  movel([-0.240083, -0.819456, -2.773882, -1.119051, 1.570796, 1.330713],accel_mss,speed_ms,0,blend_radius_m)
  movel([-0.246972, -0.827519, -2.772360, -1.112509, 1.570796, 1.323824],accel_mss,speed_ms,0,blend_radius_m)
  movel([-0.253406, -0.835845, -2.770751, -1.105793, 1.570796, 1.317390],accel_mss,speed_ms,0,blend_radius_m)
  movel([-0.259324, -0.844374, -2.769062, -1.098952, 1.570796, 1.311472],accel_mss,speed_ms,0,blend_radius_m)
  movel([-0.264353, -0.852401, -2.767435, -1.092553, 1.570796, 1.306443],accel_mss,speed_ms,0,blend_radius_m)
  movel([-0.268744, -0.860169, -2.765824, -1.086396, 1.570796, 1.302052],accel_mss,speed_ms,0,blend_radius_m)
  movel([-0.272465, -0.867667, -2.764235, -1.080487, 1.570796, 1.298331],accel_mss,speed_ms,0,blend_radius_m)
  movel([-0.275488, -0.874892, -2.762673, -1.074824, 1.570796, 1.295308],accel_mss,speed_ms,0,blend_radius_m)
  movel([-0.276730, -0.878403, -2.761902, -1.072084, 1.570796, 1.294066],accel_mss,speed_ms,0,blend_radius_m)
  movel([-0.278648, -0.885206, -2.760387, -1.066796, 1.570796, 1.292148],accel_mss,speed_ms,0,blend_radius_m)
  movel([-0.279316, -0.888500, -2.759643, -1.064245, 1.570796, 1.291480],accel_mss,speed_ms,0,blend_radius_m)
  movel([-0.280060, -0.894869, -2.758187, -1.059334, 1.570796, 1.290737],accel_mss,speed_ms,0,blend_radius_m)
  movel([-0.280127, -0.897947, -2.757473, -1.056968, 1.570796, 1.290669],accel_mss,speed_ms,0,blend_radius_m)
  movel([-0.279987, -0.900948, -2.756772, -1.054668, 1.570796, 1.290809],accel_mss,speed_ms,0,blend_radius_m)
  movel([-0.279491, -0.905065, -2.755801, -1.051523, 1.570796, 1.291305],accel_mss,speed_ms,0,blend_radius_m)
  movel([-0.278705, -0.908998, -2.754863, -1.048528, 1.570796, 1.292092],accel_mss,speed_ms,0,blend_radius_m)
  movel([-0.277654, -0.912736, -2.753962, -1.045690, 1.570796, 1.293142],accel_mss,speed_ms,0,blend_radius_m)
  movel([-0.276370, -0.916287, -2.753099, -1.043004, 1.570796, 1.294426],accel_mss,speed_ms,0,blend_radius_m)
  movel([-0.274870, -0.919629, -2.752278, -1.040482, 1.570796, 1.295926],accel_mss,speed_ms,0,blend_radius_m)
  movel([-0.273177, -0.922754, -2.751504, -1.038131, 1.570796, 1.297619],accel_mss,speed_ms,0,blend_radius_m)
  movel([-0.271316, -0.925662, -2.750778, -1.035949, 1.570796, 1.299480],accel_mss,speed_ms,0,blend_radius_m)
  movel([-0.269306, -0.928336, -2.750106, -1.033947, 1.570796, 1.301490],accel_mss,speed_ms,0,blend_radius_m)
  movel([-0.260160, -0.937511, -2.747762, -1.027116, 1.570796, 1.310636],accel_mss,speed_ms,0,blend_radius_m)
  movel([-0.253034, -0.945065, -2.745789, -1.021535, 1.570796, 1.317763],accel_mss,speed_ms,0,blend_radius_m)
  movel([-0.252477, -0.945898, -2.745569, -1.020921, 1.570796, 1.318320],accel_mss,speed_ms,0,blend_radius_m)
  movel([-0.246274, -0.937106, -2.747867, -1.027417, 1.570796, 1.324523],accel_mss,speed_ms,0,blend_radius_m)
  movel([-0.239566, -0.928371, -2.750097, -1.033921, 1.570796, 1.331230],accel_mss,speed_ms,0,blend_radius_m)
  movel([-0.232400, -0.919726, -2.752254, -1.040409, 1.570796, 1.338397],accel_mss,speed_ms,0,blend_radius_m)
  movel([-0.224833, -0.911212, -2.754331, -1.046846, 1.570796, 1.345963],accel_mss,speed_ms,0,blend_radius_m)
  movel([-0.216924, -0.902878, -2.756318, -1.053193, 1.570796, 1.353873],accel_mss,speed_ms,0,blend_radius_m)
  movel([-0.208734, -0.894762, -2.758211, -1.059416, 1.570796, 1.362062],accel_mss,speed_ms,0,blend_radius_m)
  movel([-0.200327, -0.886916, -2.760002, -1.065471, 1.570796, 1.370469],accel_mss,speed_ms,0,blend_radius_m)
  movel([-0.191774, -0.879388, -2.761684, -1.071317, 1.570796, 1.379022],accel_mss,speed_ms,0,blend_radius_m)
  movel([-0.187679, -0.876001, -2.762430, -1.073958, 1.570796, 1.383118],accel_mss,speed_ms,0,blend_radius_m)
  movel([-0.183450, -0.872734, -2.763143, -1.076512, 1.570796, 1.387346],accel_mss,speed_ms,0,blend_radius_m)
  movel([-0.179125, -0.869625, -2.763815, -1.078949, 1.570796, 1.391671],accel_mss,speed_ms,0,blend_radius_m)
  movel([-0.174747, -0.866715, -2.764439, -1.081235, 1.570796, 1.396049],accel_mss,speed_ms,0,blend_radius_m)
  movel([-0.170354, -0.864043, -2.765007, -1.083339, 1.570796, 1.400443],accel_mss,speed_ms,0,blend_radius_m)
  movel([-0.165982, -0.861648, -2.765513, -1.085228, 1.570796, 1.404814],accel_mss,speed_ms,0,blend_radius_m)
  movel([-0.161676, -0.859568, -2.765950, -1.086871, 1.570796, 1.409121],accel_mss,speed_ms,0,blend_radius_m)
  movel([-0.157477, -0.857842, -2.766310, -1.088237, 1.570796, 1.413319],accel_mss,speed_ms,0,blend_radius_m)
  movel([-0.153425, -0.856510, -2.766587, -1.089292, 1.570796, 1.417371],accel_mss,speed_ms,0,blend_radius_m)
  movel([-0.149560, -0.855608, -2.766774, -1.090007, 1.570796, 1.421237],accel_mss,speed_ms,0,blend_radius_m)
  movel([-0.145927, -0.855177, -2.766863, -1.090349, 1.570796, 1.424869],accel_mss,speed_ms,0,blend_radius_m)
  movel([-0.142567, -0.855251, -2.766848, -1.090290, 1.570796, 1.428229],accel_mss,speed_ms,0,blend_radius_m)
  movel([-0.139522, -0.855865, -2.766721, -1.089803, 1.570796, 1.431274],accel_mss,speed_ms,0,blend_radius_m)
  movel([-0.136824, -0.857050, -2.766475, -1.088864, 1.570796, 1.433972],accel_mss,speed_ms,0,blend_radius_m)
  movel([-0.134519, -0.858837, -2.766102, -1.087449, 1.570796, 1.436278],accel_mss,speed_ms,0,blend_radius_m)
  movel([-0.132645, -0.861261, -2.765595, -1.085534, 1.570796, 1.438152],accel_mss,speed_ms,0,blend_radius_m)
  movel([-0.130842, -0.865165, -2.764769, -1.082455, 1.570796, 1.439954],accel_mss,speed_ms,0,blend_radius_m)
  movel([-0.129631, -0.869711, -2.763796, -1.078881, 1.570796, 1.441165],accel_mss,speed_ms,0,blend_radius_m)
  movel([-0.128936, -0.874759, -2.762702, -1.074928, 1.570796, 1.441860],accel_mss,speed_ms,0,blend_radius_m)
  movel([-0.128670, -0.880175, -2.761510, -1.070704, 1.570796, 1.442126],accel_mss,speed_ms,0,blend_radius_m)
  movel([-0.128760, -0.885825, -2.760248, -1.066316, 1.570796, 1.442036],accel_mss,speed_ms,0,blend_radius_m)
  movel([-0.129131, -0.891586, -2.758941, -1.061862, 1.570796, 1.441665],accel_mss,speed_ms,0,blend_radius_m)
  movel([-0.130394, -0.902931, -2.756306, -1.053152, 1.570796, 1.440402],accel_mss,speed_ms,0,blend_radius_m)
  movel([-0.131557, -0.910187, -2.754578, -1.047624, 1.570796, 1.439239],accel_mss,speed_ms,0,blend_radius_m)
  movel([-0.133085, -0.917458, -2.752812, -1.042119, 1.570796, 1.437712],accel_mss,speed_ms,0,blend_radius_m)
  movel([-0.134926, -0.924737, -2.751010, -1.036643, 1.570796, 1.435870],accel_mss,speed_ms,0,blend_radius_m)
  movel([-0.137037, -0.932034, -2.749168, -1.031187, 1.570796, 1.433760],accel_mss,speed_ms,0,blend_radius_m)
  movel([-0.139370, -0.939343, -2.747287, -1.025759, 1.570796, 1.431427],accel_mss,speed_ms,0,blend_radius_m)
  movel([-0.141879, -0.946667, -2.745366, -1.020356, 1.570796, 1.428917],accel_mss,speed_ms,0,blend_radius_m)
  movel([-0.147269, -0.961389, -2.741392, -1.009608, 1.570796, 1.423527],accel_mss,speed_ms,0,blend_radius_m)
  movel([-0.140519, -0.960936, -2.741517, -1.009936, 1.570796, 1.430278],accel_mss,speed_ms,0,blend_radius_m)
  movel([-0.137016, -0.960927, -2.741519, -1.009943, 1.570796, 1.433781],accel_mss,speed_ms,0,blend_radius_m)
  movel([-0.133979, -0.961411, -2.741386, -1.009592, 1.570796, 1.436818],accel_mss,speed_ms,0,blend_radius_m)
  movel([-0.132765, -0.961921, -2.741245, -1.009222, 1.570796, 1.438031],accel_mss,speed_ms,0,blend_radius_m)
  movel([-0.131825, -0.962655, -2.741043, -1.008690, 1.570796, 1.438971],accel_mss,speed_ms,0,blend_radius_m)
  movel([-0.131206, -0.963639, -2.740771, -1.007979, 1.570796, 1.439590],accel_mss,speed_ms,0,blend_radius_m)
  movel([-0.130958, -0.964905, -2.740420, -1.007064, 1.570796, 1.439839],accel_mss,speed_ms,0,blend_radius_m)
  movel([-0.131131, -0.966478, -2.739983, -1.005928, 1.570796, 1.439665],accel_mss,speed_ms,0,blend_radius_m)
  movel([-0.131778, -0.968398, -2.739446, -1.004544, 1.570796, 1.439018],accel_mss,speed_ms,0,blend_radius_m)
  movel([-0.132943, -0.970690, -2.738802, -1.002896, 1.570796, 1.437853],accel_mss,speed_ms,0,blend_radius_m)
  movel([-0.134674, -0.973378, -2.738043, -1.000969, 1.570796, 1.436123],accel_mss,speed_ms,0,blend_radius_m)
  movel([-0.136314, -0.975590, -2.737413, -0.999386, 1.570796, 1.434482],accel_mss,speed_ms,0,blend_radius_m)
  movel([-0.137990, -0.977600, -2.736838, -0.997950, 1.570796, 1.432806],accel_mss,speed_ms,0,blend_radius_m)
  movel([-0.139696, -0.979424, -2.736314, -0.996651, 1.570796, 1.431100],accel_mss,speed_ms,0,blend_radius_m)
  movel([-0.143196, -0.982582, -2.735401, -0.994406, 1.570796, 1.427601],accel_mss,speed_ms,0,blend_radius_m)
  movel([-0.144982, -0.983947, -2.735004, -0.993438, 1.570796, 1.425815],accel_mss,speed_ms,0,blend_radius_m)
  movel([-0.148619, -0.986335, -2.734306, -0.991748, 1.570796, 1.422177],accel_mss,speed_ms,0,blend_radius_m)
  movel([-0.152315, -0.988361, -2.733710, -0.990318, 1.570796, 1.418481],accel_mss,speed_ms,0,blend_radius_m)
  movel([-0.156050, -0.990151, -2.733182, -0.989056, 1.570796, 1.414746],accel_mss,speed_ms,0,blend_radius_m)
  movel([-0.163527, -0.993487, -2.732190, -0.986712, 1.570796, 1.407269],accel_mss,speed_ms,0,blend_radius_m)
  movel([-0.166909, -0.999532, -2.730372, -0.982486, 1.570796, 1.403888],accel_mss,speed_ms,0,blend_radius_m)
  movel([-0.168793, -1.002571, -2.729447, -0.980371, 1.570796, 1.402004],accel_mss,speed_ms,0,blend_radius_m)
  movel([-0.170824, -1.005546, -2.728535, -0.978308, 1.570796, 1.399972],accel_mss,speed_ms,0,blend_radius_m)
  movel([-0.173015, -1.008396, -2.727655, -0.976338, 1.570796, 1.397781],accel_mss,speed_ms,0,blend_radius_m)
  movel([-0.175376, -1.011062, -2.726826, -0.974501, 1.570796, 1.395420],accel_mss,speed_ms,0,blend_radius_m)
  movel([-0.177921, -1.013486, -2.726068, -0.972835, 1.570796, 1.392875],accel_mss,speed_ms,0,blend_radius_m)
  movel([-0.180668, -1.015618, -2.725397, -0.971375, 1.570796, 1.390128],accel_mss,speed_ms,0,blend_radius_m)
  movel([-0.182641, -1.016748, -2.725040, -0.970601, 1.570796, 1.388155],accel_mss,speed_ms,0,blend_radius_m)
  movel([-0.184252, -1.017225, -2.724889, -0.970275, 1.570796, 1.386545],accel_mss,speed_ms,0,blend_radius_m)
  movel([-0.185536, -1.017141, -2.724915, -0.970332, 1.570796, 1.385261],accel_mss,speed_ms,0,blend_radius_m)
  movel([-0.186525, -1.016588, -2.725090, -0.970711, 1.570796, 1.384271],accel_mss,speed_ms,0,blend_radius_m)
  movel([-0.187255, -1.015653, -2.725386, -0.971350, 1.570796, 1.383541],accel_mss,speed_ms,0,blend_radius_m)
  movel([-0.187753, -1.014434, -2.725770, -0.972185, 1.570796, 1.383044],accel_mss,speed_ms,0,blend_radius_m)
  movel([-0.188056, -1.013020, -2.726214, -0.973155, 1.570796, 1.382740],accel_mss,speed_ms,0,blend_radius_m)
  movel([-0.188187, -1.011496, -2.726691, -0.974202, 1.570796, 1.382610],accel_mss,speed_ms,0,blend_radius_m)
  movel([-0.188105, -1.008082, -2.727752, -0.976554, 1.570796, 1.382691],accel_mss,speed_ms,0,blend_radius_m)
  movel([-0.187675, -1.004518, -2.728851, -0.979020, 1.570796, 1.383122],accel_mss,speed_ms,0,blend_radius_m)
  movel([-0.186308, -0.997047, -2.731122, -0.984220, 1.570796, 1.384488],accel_mss,speed_ms,0,blend_radius_m)
  movel([-0.195311, -0.996681, -2.731233, -0.984476, 1.570796, 1.375486],accel_mss,speed_ms,0,blend_radius_m)
  movel([-0.204501, -0.996669, -2.731236, -0.984483, 1.570796, 1.366295],accel_mss,speed_ms,0,blend_radius_m)
  movel([-0.213681, -0.996628, -2.731248, -0.984512, 1.570796, 1.357115],accel_mss,speed_ms,0,blend_radius_m)
  movel([-0.218210, -0.996477, -2.731294, -0.984618, 1.570796, 1.352586],accel_mss,speed_ms,0,blend_radius_m)
  movel([-0.222670, -0.996174, -2.731385, -0.984830, 1.570796, 1.348127],accel_mss,speed_ms,0,blend_radius_m)
  movel([-0.226835, -0.995688, -2.731531, -0.985170, 1.570796, 1.343961],accel_mss,speed_ms,0,blend_radius_m)
  movel([-0.230874, -0.995032, -2.731728, -0.985630, 1.570796, 1.339922],accel_mss,speed_ms,0,blend_radius_m)
  movel([-0.238718, -0.993394, -2.732218, -0.986777, 1.570796, 1.332079],accel_mss,speed_ms,0,blend_radius_m)
  movel([-0.246507, -0.991697, -2.732723, -0.987969, 1.570796, 1.324289],accel_mss,speed_ms,0,blend_radius_m)
  movel([-0.254533, -0.990366, -2.733118, -0.988905, 1.570796, 1.316263],accel_mss,speed_ms,0,blend_radius_m)
  movel([-0.255753, -0.994675, -2.731835, -0.985880, 1.570796, 1.315043],accel_mss,speed_ms,0,blend_radius_m)
  movel([-0.256733, -0.998854, -2.730577, -0.982958, 1.570796, 1.314063],accel_mss,speed_ms,0,blend_radius_m)
  movel([-0.257476, -1.002898, -2.729347, -0.980144, 1.570796, 1.313321],accel_mss,speed_ms,0,blend_radius_m)
  movel([-0.257986, -1.006800, -2.728149, -0.977441, 1.570796, 1.312810],accel_mss,speed_ms,0,blend_radius_m)
  movel([-0.258266, -1.010558, -2.726983, -0.974848, 1.570796, 1.312531],accel_mss,speed_ms,0,blend_radius_m)
  movel([-0.258324, -1.014167, -2.725854, -0.972368, 1.570796, 1.312472],accel_mss,speed_ms,0,blend_radius_m)
  movel([-0.258158, -1.017623, -2.724762, -0.970003, 1.570796, 1.312639],accel_mss,speed_ms,0,blend_radius_m)
  movel([-0.257779, -1.020927, -2.723711, -0.967751, 1.570796, 1.313017],accel_mss,speed_ms,0,blend_radius_m)
  movel([-0.257186, -1.024070, -2.722702, -0.965617, 1.570796, 1.313610],accel_mss,speed_ms,0,blend_radius_m)
  movel([-0.256379, -1.027045, -2.721740, -0.963604, 1.570796, 1.314417],accel_mss,speed_ms,0,blend_radius_m)
  movel([-0.255369, -1.029859, -2.720824, -0.961707, 1.570796, 1.315428],accel_mss,speed_ms,0,blend_radius_m)
  movel([-0.254157, -1.032501, -2.719957, -0.959931, 1.570796, 1.316640],accel_mss,speed_ms,0,blend_radius_m)
  movel([-0.252740, -1.034963, -2.719145, -0.958281, 1.570796, 1.318057],accel_mss,speed_ms,0,blend_radius_m)
  movel([-0.251127, -1.037252, -2.718385, -0.956752, 1.570796, 1.319670],accel_mss,speed_ms,0,blend_radius_m)
  movel([-0.249319, -1.039357, -2.717683, -0.955349, 1.570796, 1.321477],accel_mss,speed_ms,0,blend_radius_m)
  movel([-0.247315, -1.041276, -2.717039, -0.954073, 1.570796, 1.323481],accel_mss,speed_ms,0,blend_radius_m)
  movel([-0.243873, -1.043875, -2.716163, -0.952351, 1.570796, 1.326923],accel_mss,speed_ms,0,blend_radius_m)
  movel([-0.240108, -1.046022, -2.715435, -0.950932, 1.570796, 1.330689],accel_mss,speed_ms,0,blend_radius_m)
  movel([-0.236060, -1.047768, -2.714840, -0.949781, 1.570796, 1.334737],accel_mss,speed_ms,0,blend_radius_m)
  movel([-0.231757, -1.049149, -2.714368, -0.948872, 1.570796, 1.339039],accel_mss,speed_ms,0,blend_radius_m)
  movel([-0.227241, -1.050211, -2.714003, -0.948174, 1.570796, 1.343555],accel_mss,speed_ms,0,blend_radius_m)
  movel([-0.222546, -1.050993, -2.713735, -0.947661, 1.570796, 1.348251],accel_mss,speed_ms,0,blend_radius_m)
  movel([-0.217707, -1.051537, -2.713547, -0.947304, 1.570796, 1.353089],accel_mss,speed_ms,0,blend_radius_m)
  movel([-0.212754, -1.051872, -2.713432, -0.947085, 1.570796, 1.358042],accel_mss,speed_ms,0,blend_radius_m)
  movel([-0.202592, -1.052132, -2.713342, -0.946915, 1.570796, 1.368205],accel_mss,speed_ms,0,blend_radius_m)
  movel([-0.192313, -1.052163, -2.713332, -0.946895, 1.570796, 1.378484],accel_mss,speed_ms,0,blend_radius_m)
  movel([-0.184486, -1.052432, -2.713239, -0.946719, 1.570796, 1.386310],accel_mss,speed_ms,0,blend_radius_m)
  movel([-0.181810, -1.052339, -2.713271, -0.946779, 1.570796, 1.388986],accel_mss,speed_ms,0,blend_radius_m)
  movel([-0.177019, -1.051809, -2.713454, -0.947126, 1.570796, 1.393777],accel_mss,speed_ms,0,blend_radius_m)
  movel([-0.176000, -1.051875, -2.713431, -0.947083, 1.570796, 1.394796],accel_mss,speed_ms,0,blend_radius_m)
  movel([-0.175063, -1.052126, -2.713344, -0.946919, 1.570796, 1.395734],accel_mss,speed_ms,0,blend_radius_m)
  movel([-0.174219, -1.052622, -2.713173, -0.946594, 1.570796, 1.396577],accel_mss,speed_ms,0,blend_radius_m)
  movel([-0.173481, -1.053421, -2.712897, -0.946072, 1.570796, 1.397315],accel_mss,speed_ms,0,blend_radius_m)
  movel([-0.172877, -1.054584, -2.712494, -0.945312, 1.570796, 1.397920],accel_mss,speed_ms,0,blend_radius_m)
  movel([-0.172560, -1.055937, -2.712023, -0.944429, 1.570796, 1.398237],accel_mss,speed_ms,0,blend_radius_m)
  movel([-0.172504, -1.057446, -2.711496, -0.943446, 1.570796, 1.398292],accel_mss,speed_ms,0,blend_radius_m)
  movel([-0.172688, -1.059097, -2.710918, -0.942374, 1.570796, 1.398108],accel_mss,speed_ms,0,blend_radius_m)
  movel([-0.173088, -1.060854, -2.710300, -0.941235, 1.570796, 1.397708],accel_mss,speed_ms,0,blend_radius_m)
  movel([-0.174448, -1.064617, -2.708968, -0.938804, 1.570796, 1.396348],accel_mss,speed_ms,0,blend_radius_m)
  movel([-0.175364, -1.066571, -2.708271, -0.937547, 1.570796, 1.395432],accel_mss,speed_ms,0,blend_radius_m)
  movel([-0.177543, -1.070508, -2.706857, -0.935024, 1.570796, 1.393253],accel_mss,speed_ms,0,blend_radius_m)
  movel([-0.180056, -1.074338, -2.705469, -0.932582, 1.570796, 1.390741],accel_mss,speed_ms,0,blend_radius_m)
  movel([-0.182720, -1.077881, -2.704173, -0.930334, 1.570796, 1.388077],accel_mss,speed_ms,0,blend_radius_m)
  movel([-0.185375, -1.080971, -2.703035, -0.928384, 1.570796, 1.385422],accel_mss,speed_ms,0,blend_radius_m)
  movel([-0.189597, -1.085203, -2.701461, -0.925725, 1.570796, 1.381199],accel_mss,speed_ms,0,blend_radius_m)
  movel([-0.191807, -1.087186, -2.700718, -0.924485, 1.570796, 1.378989],accel_mss,speed_ms,0,blend_radius_m)
  movel([-0.194067, -1.089067, -2.700010, -0.923312, 1.570796, 1.376730],accel_mss,speed_ms,0,blend_radius_m)
  movel([-0.198705, -1.092523, -2.698702, -0.921165, 1.570796, 1.372091],accel_mss,speed_ms,0,blend_radius_m)
  movel([-0.203436, -1.095533, -2.697553, -0.919303, 1.570796, 1.367360],accel_mss,speed_ms,0,blend_radius_m)
  movel([-0.208189, -1.098060, -2.696582, -0.917747, 1.570796, 1.362608],accel_mss,speed_ms,0,blend_radius_m)
  movel([-0.212880, -1.100063, -2.695808, -0.916517, 1.570796, 1.357916],accel_mss,speed_ms,0,blend_radius_m)
  movel([-0.215184, -1.100855, -2.695502, -0.916032, 1.570796, 1.355612],accel_mss,speed_ms,0,blend_radius_m)
  movel([-0.219661, -1.101997, -2.695058, -0.915334, 1.570796, 1.351136],accel_mss,speed_ms,0,blend_radius_m)
  movel([-0.221816, -1.102335, -2.694927, -0.915128, 1.570796, 1.348981],accel_mss,speed_ms,0,blend_radius_m)
  movel([-0.224573, -1.102550, -2.694843, -0.914996, 1.570796, 1.346223],accel_mss,speed_ms,0,blend_radius_m)
  movel([-0.227217, -1.102535, -2.694849, -0.915005, 1.570796, 1.343579],accel_mss,speed_ms,0,blend_radius_m)
  movel([-0.229757, -1.102317, -2.694933, -0.915138, 1.570796, 1.341039],accel_mss,speed_ms,0,blend_radius_m)
  movel([-0.232211, -1.101933, -2.695083, -0.915373, 1.570796, 1.338585],accel_mss,speed_ms,0,blend_radius_m)
  movel([-0.236912, -1.100784, -2.695529, -0.916076, 1.570796, 1.333885],accel_mss,speed_ms,0,blend_radius_m)
  movel([-0.241425, -1.099339, -2.696089, -0.916962, 1.570796, 1.329371],accel_mss,speed_ms,0,blend_radius_m)
  movel([-0.246938, -1.097314, -2.696869, -0.918206, 1.570796, 1.323859],accel_mss,speed_ms,0,blend_radius_m)
  movel([-0.252299, -1.095002, -2.697756, -0.919631, 1.570796, 1.318497],accel_mss,speed_ms,0,blend_radius_m)
  movel([-0.257469, -1.092384, -2.698754, -0.921251, 1.570796, 1.313328],accel_mss,speed_ms,0,blend_radius_m)
  movel([-0.262410, -1.089440, -2.699870, -0.923079, 1.570796, 1.308386],accel_mss,speed_ms,0,blend_radius_m)
  movel([-0.267082, -1.086144, -2.701109, -0.925136, 1.570796, 1.303714],accel_mss,speed_ms,0,blend_radius_m)
  movel([-0.271439, -1.082471, -2.702479, -0.927439, 1.570796, 1.299357],accel_mss,speed_ms,0,blend_radius_m)
  movel([-0.275442, -1.078397, -2.703984, -0.930008, 1.570796, 1.295354],accel_mss,speed_ms,0,blend_radius_m)
  movel([-0.279047, -1.073894, -2.705631, -0.932864, 1.570796, 1.291750],accel_mss,speed_ms,0,blend_radius_m)
  movel([-0.281489, -1.070225, -2.706959, -0.935205, 1.570796, 1.289307],accel_mss,speed_ms,0,blend_radius_m)
  movel([-0.283792, -1.066194, -2.708406, -0.937789, 1.570796, 1.287004],accel_mss,speed_ms,0,blend_radius_m)
  movel([-0.285884, -1.061819, -2.709960, -0.940611, 1.570796, 1.284912],accel_mss,speed_ms,0,blend_radius_m)
  movel([-0.287694, -1.057127, -2.711608, -0.943654, 1.570796, 1.283102],accel_mss,speed_ms,0,blend_radius_m)
  movel([-0.289143, -1.052140, -2.713340, -0.946910, 1.570796, 1.281653],accel_mss,speed_ms,0,blend_radius_m)
  movel([-0.290151, -1.046878, -2.715144, -0.950367, 1.570796, 1.280645],accel_mss,speed_ms,0,blend_radius_m)
  movel([-0.290644, -1.041362, -2.717011, -0.954017, 1.570796, 1.280153],accel_mss,speed_ms,0,blend_radius_m)
  movel([-0.290668, -1.038512, -2.717965, -0.955912, 1.570796, 1.280128],accel_mss,speed_ms,0,blend_radius_m)
  movel([-0.290533, -1.035608, -2.718931, -0.957850, 1.570796, 1.280264],accel_mss,speed_ms,0,blend_radius_m)
  movel([-0.289916, -1.029983, -2.720783, -0.961623, 1.570796, 1.280881],accel_mss,speed_ms,0,blend_radius_m)
  movel([-0.288898, -1.024139, -2.722680, -0.965570, 1.570796, 1.281898],accel_mss,speed_ms,0,blend_radius_m)
  movel([-0.287475, -1.018094, -2.724613, -0.969682, 1.570796, 1.283321],accel_mss,speed_ms,0,blend_radius_m)
  movel([-0.285657, -1.011872, -2.726573, -0.973944, 1.570796, 1.285140],accel_mss,speed_ms,0,blend_radius_m)
  movel([-0.283430, -1.005489, -2.728552, -0.978347, 1.570796, 1.287366],accel_mss,speed_ms,0,blend_radius_m)
  movel([-0.280808, -0.998974, -2.730540, -0.982874, 1.570796, 1.289988],accel_mss,speed_ms,0,blend_radius_m)
  movel([-0.277785, -0.992346, -2.732530, -0.987513, 1.570796, 1.293011],accel_mss,speed_ms,0,blend_radius_m)
  movel([-0.274360, -0.985633, -2.734511, -0.992245, 1.570796, 1.296436],accel_mss,speed_ms,0,blend_radius_m)
  movel([-0.284136, -0.979906, -2.736175, -0.996308, 1.570796, 1.286660],accel_mss,speed_ms,0,blend_radius_m)
  movel([-0.289076, -0.977084, -2.736986, -0.998319, 1.570796, 1.281720],accel_mss,speed_ms,0,blend_radius_m)
  movel([-0.293829, -0.973999, -2.737866, -1.000524, 1.570796, 1.276967],accel_mss,speed_ms,0,blend_radius_m)
  movel([-0.297075, -0.971319, -2.738625, -1.002445, 1.570796, 1.273721],accel_mss,speed_ms,0,blend_radius_m)
  movel([-0.299951, -0.968195, -2.739503, -1.004691, 1.570796, 1.270845],accel_mss,speed_ms,0,blend_radius_m)
  movel([-0.302469, -0.964659, -2.740489, -1.007241, 1.570796, 1.268328],accel_mss,speed_ms,0,blend_radius_m)
  movel([-0.304635, -0.960728, -2.741574, -1.010087, 1.570796, 1.266162],accel_mss,speed_ms,0,blend_radius_m)
  movel([-0.306456, -0.956428, -2.742748, -1.013213, 1.570796, 1.264341],accel_mss,speed_ms,0,blend_radius_m)
  movel([-0.307936, -0.951780, -2.744003, -1.016606, 1.570796, 1.262860],accel_mss,speed_ms,0,blend_radius_m)
  movel([-0.309084, -0.946806, -2.745329, -1.020254, 1.570796, 1.261712],accel_mss,speed_ms,0,blend_radius_m)
  movel([-0.309905, -0.941531, -2.746717, -1.024141, 1.570796, 1.260892],accel_mss,speed_ms,0,blend_radius_m)
  movel([-0.310400, -0.935981, -2.748156, -1.028251, 1.570796, 1.260397],accel_mss,speed_ms,0,blend_radius_m)
  movel([-0.310573, -0.930172, -2.749641, -1.032576, 1.570796, 1.260223],accel_mss,speed_ms,0,blend_radius_m)
  movel([-0.310429, -0.924132, -2.751161, -1.037097, 1.570796, 1.260367],accel_mss,speed_ms,0,blend_radius_m)
  movel([-0.309975, -0.917888, -2.752707, -1.041795, 1.570796, 1.260822],accel_mss,speed_ms,0,blend_radius_m)
  movel([-0.309210, -0.911464, -2.754270, -1.046655, 1.570796, 1.261586],accel_mss,speed_ms,0,blend_radius_m)
  movel([-0.308145, -0.904896, -2.755841, -1.051652, 1.570796, 1.262651],accel_mss,speed_ms,0,blend_radius_m)
  movel([-0.306775, -0.898199, -2.757415, -1.056775, 1.570796, 1.264021],accel_mss,speed_ms,0,blend_radius_m)
  movel([-0.305113, -0.891413, -2.758980, -1.061996, 1.570796, 1.265683],accel_mss,speed_ms,0,blend_radius_m)
  movel([-0.301396, -0.878383, -2.761906, -1.072100, 1.570796, 1.269401],accel_mss,speed_ms,0,blend_radius_m)
  movel([-0.299215, -0.871668, -2.763374, -1.077347, 1.570796, 1.271582],accel_mss,speed_ms,0,blend_radius_m)
  movel([-0.296761, -0.864817, -2.764843, -1.082729, 1.570796, 1.274035],accel_mss,speed_ms,0,blend_radius_m)
  movel([-0.293979, -0.857832, -2.766312, -1.088245, 1.570796, 1.276817],accel_mss,speed_ms,0,blend_radius_m)
  movel([-0.290827, -0.850719, -2.767779, -1.093891, 1.570796, 1.279970],accel_mss,speed_ms,0,blend_radius_m)
  movel([-0.287253, -0.843476, -2.769242, -1.099671, 1.570796, 1.283543],accel_mss,speed_ms,0,blend_radius_m)
  movel([-0.283205, -0.836106, -2.770700, -1.105583, 1.570796, 1.287592],accel_mss,speed_ms,0,blend_radius_m)
  movel([-0.278188, -0.827816, -2.772304, -1.112269, 1.570796, 1.292608],accel_mss,speed_ms,0,blend_radius_m)
  movel([-0.272701, -0.819458, -2.773882, -1.119049, 1.570796, 1.298096],accel_mss,speed_ms,0,blend_radius_m)
  movel([-0.266775, -0.811057, -2.775429, -1.125903, 1.570796, 1.304021],accel_mss,speed_ms,0,blend_radius_m)
  movel([-0.260437, -0.802648, -2.776939, -1.132802, 1.570796, 1.310359],accel_mss,speed_ms,0,blend_radius_m)
  movel([-0.253721, -0.794265, -2.778407, -1.139717, 1.570796, 1.317075],accel_mss,speed_ms,0,blend_radius_m)
  movel([-0.246662, -0.785948, -2.779827, -1.146614, 1.570796, 1.324135],accel_mss,speed_ms,0,blend_radius_m)
  movel([-0.239288, -0.777726, -2.781196, -1.153467, 1.570796, 1.331508],accel_mss,speed_ms,0,blend_radius_m)
  movel([-0.231644, -0.769647, -2.782506, -1.160236, 1.570796, 1.339152],accel_mss,speed_ms,0,blend_radius_m)
  movel([-0.223767, -0.761753, -2.783755, -1.166881, 1.570796, 1.347029],accel_mss,speed_ms,0,blend_radius_m)
  movel([-0.215708, -0.754085, -2.784938, -1.173365, 1.570796, 1.355088],accel_mss,speed_ms,0,blend_radius_m)
  movel([-0.207502, -0.746689, -2.786052, -1.179648, 1.570796, 1.363295],accel_mss,speed_ms,0,blend_radius_m)
  movel([-0.199198, -0.739607, -2.787093, -1.185689, 1.570796, 1.371598],accel_mss,speed_ms,0,blend_radius_m)
  movel([-0.190853, -0.732893, -2.788058, -1.191438, 1.570796, 1.379943],accel_mss,speed_ms,0,blend_radius_m)
  movel([-0.182509, -0.726584, -2.788945, -1.196860, 1.570796, 1.388287],accel_mss,speed_ms,0,blend_radius_m)
  movel([-0.174221, -0.720731, -2.789751, -1.201907, 1.570796, 1.396576],accel_mss,speed_ms,0,blend_radius_m)
  movel([-0.166037, -0.715380, -2.790473, -1.206536, 1.570796, 1.404759],accel_mss,speed_ms,0,blend_radius_m)
  movel([-0.157405, -0.710096, -2.791174, -1.211119, 1.570796, 1.413391],accel_mss,speed_ms,0,blend_radius_m)
  movel([-0.148804, -0.705148, -2.791818, -1.215423, 1.570796, 1.421992],accel_mss,speed_ms,0,blend_radius_m)
  movel([-0.140291, -0.700650, -2.792394, -1.219345, 1.570796, 1.430505],accel_mss,speed_ms,0,blend_radius_m)
  movel([-0.131927, -0.696734, -2.792888, -1.222767, 1.570796, 1.438870],accel_mss,speed_ms,0,blend_radius_m)
  movel([-0.122400, -0.693002, -2.793352, -1.226035, 1.570796, 1.448396],accel_mss,speed_ms,0,blend_radius_m)
  movel([-0.113109, -0.690149, -2.793703, -1.228538, 1.570796, 1.457687],accel_mss,speed_ms,0,blend_radius_m)
  movel([-0.104162, -0.688206, -2.793939, -1.230244, 1.570796, 1.466634],accel_mss,speed_ms,0,blend_radius_m)
  movel([-0.095662, -0.687199, -2.794061, -1.231129, 1.570796, 1.475134],accel_mss,speed_ms,0,blend_radius_m)
  movel([-0.087705, -0.687142, -2.794068, -1.231179, 1.570796, 1.483091],accel_mss,speed_ms,0,blend_radius_m)
  movel([-0.080386, -0.688045, -2.793959, -1.230385, 1.570796, 1.490410],accel_mss,speed_ms,0,blend_radius_m)
  movel([-0.073790, -0.689903, -2.793733, -1.228753, 1.570796, 1.497006],accel_mss,speed_ms,0,blend_radius_m)
  movel([-0.067994, -0.692714, -2.793388, -1.226288, 1.570796, 1.502802],accel_mss,speed_ms,0,blend_radius_m)
  movel([-0.057560, -0.699516, -2.792538, -1.220335, 1.570796, 1.513236],accel_mss,speed_ms,0,blend_radius_m)
  movel([-0.052798, -0.703410, -2.792042, -1.216937, 1.570796, 1.517998],accel_mss,speed_ms,0,blend_radius_m)
  movel([-0.048479, -0.707967, -2.791452, -1.212969, 1.570796, 1.522318],accel_mss,speed_ms,0,blend_radius_m)
  movel([-0.041507, -0.715992, -2.790391, -1.206006, 1.570796, 1.529289],accel_mss,speed_ms,0,blend_radius_m)
  movel([-0.037675, -0.719700, -2.789891, -1.202798, 1.570796, 1.533121],accel_mss,speed_ms,0,blend_radius_m)
  movel([-0.033523, -0.723005, -2.789439, -1.199945, 1.570796, 1.537274],accel_mss,speed_ms,0,blend_radius_m)
  movel([-0.028962, -0.725750, -2.789061, -1.197579, 1.570796, 1.541834],accel_mss,speed_ms,0,blend_radius_m)
  movel([-0.023934, -0.727791, -2.788777, -1.195821, 1.570796, 1.546863],accel_mss,speed_ms,0,blend_radius_m)
  movel([-0.018345, -0.728973, -2.788611, -1.194805, 1.570796, 1.552452],accel_mss,speed_ms,0,blend_radius_m)
  movel([-0.012124, -0.729146, -2.788587, -1.194656, 1.570796, 1.558673],accel_mss,speed_ms,0,blend_radius_m)
  movel([-0.009390, -0.728804, -2.788635, -1.194950, 1.570796, 1.561406],accel_mss,speed_ms,0,blend_radius_m)
  movel([-0.006411, -0.727933, -2.788757, -1.195699, 1.570796, 1.564385],accel_mss,speed_ms,0,blend_radius_m)
  movel([-0.004852, -0.727224, -2.788856, -1.196310, 1.570796, 1.565945],accel_mss,speed_ms,0,blend_radius_m)
  movel([-0.003262, -0.726299, -2.788984, -1.197106, 1.570796, 1.567535],accel_mss,speed_ms,0,blend_radius_m)
  movel([-0.001645, -0.725127, -2.789147, -1.198115, 1.570796, 1.569152],accel_mss,speed_ms,0,blend_radius_m)
  movel([-0.000021, -0.723676, -2.789347, -1.199365, 1.570796, 1.570776],accel_mss,speed_ms,0,blend_radius_m)
  movel([0.001581, -0.721953, -2.789584, -1.200852, 1.570796, 1.572377],accel_mss,speed_ms,0,blend_radius_m)
  movel([0.003048, -0.720085, -2.789839, -1.202465, 1.570796, 1.573844],accel_mss,speed_ms,0,blend_radius_m)
  movel([0.005585, -0.716143, -2.790371, -1.205875, 1.570796, 1.576381],accel_mss,speed_ms,0,blend_radius_m)
  movel([0.007057, -0.713381, -2.790740, -1.208268, 1.570796, 1.577853],accel_mss,speed_ms,0,blend_radius_m)
  movel([0.008285, -0.710687, -2.791096, -1.210606, 1.570796, 1.579082],accel_mss,speed_ms,0,blend_radius_m)
  movel([0.010077, -0.705512, -2.791771, -1.215106, 1.570796, 1.580873],accel_mss,speed_ms,0,blend_radius_m)
  movel([0.011073, -0.700649, -2.792394, -1.219346, 1.570796, 1.581869],accel_mss,speed_ms,0,blend_radius_m)
  movel([0.011397, -0.696110, -2.792966, -1.223313, 1.570796, 1.582193],accel_mss,speed_ms,0,blend_radius_m)
  movel([0.011166, -0.691929, -2.793484, -1.226976, 1.570796, 1.581962],accel_mss,speed_ms,0,blend_radius_m)
  movel([0.010505, -0.688120, -2.793950, -1.230319, 1.570796, 1.581301],accel_mss,speed_ms,0,blend_radius_m)
  movel([0.009538, -0.684705, -2.794361, -1.233323, 1.570796, 1.580334],accel_mss,speed_ms,0,blend_radius_m)
  movel([0.006816, -0.678599, -2.795085, -1.238705, 1.570796, 1.577613],accel_mss,speed_ms,0,blend_radius_m)
  movel([0.004888, -0.675865, -2.795403, -1.241121, 1.570796, 1.575684],accel_mss,speed_ms,0,blend_radius_m)
  movel([0.002618, -0.673509, -2.795675, -1.243205, 1.570796, 1.573414],accel_mss,speed_ms,0,blend_radius_m)
  movel([0.000011, -0.671558, -2.795898, -1.244933, 1.570796, 1.570807],accel_mss,speed_ms,0,blend_radius_m)
  movel([-0.002929, -0.670023, -2.796072, -1.246293, 1.570796, 1.567867],accel_mss,speed_ms,0,blend_radius_m)
  movel([-0.006191, -0.668925, -2.796197, -1.247267, 1.570796, 1.564605],accel_mss,speed_ms,0,blend_radius_m)
  movel([-0.009757, -0.668268, -2.796271, -1.247851, 1.570796, 1.561039],accel_mss,speed_ms,0,blend_radius_m)
  movel([-0.013626, -0.668070, -2.796293, -1.248026, 1.570796, 1.557171],accel_mss,speed_ms,0,blend_radius_m)
  speed_ms = 0.005
  movel([-0.013626, -0.662122, -2.789593, -1.260673, 1.570796, 1.557171],accel_mss,speed_ms,0,blend_radius_m)
  speed_ms = 0.040
  movel([-0.011127, -0.692738, -2.785956, -1.233695, 1.570796, 1.559669],accel_mss,speed_ms,0,blend_radius_m)
  speed_ms = 0.005
  movel([-0.011127, -0.699112, -2.792589, -1.220688, 1.570796, 1.559669],accel_mss,speed_ms,0,blend_radius_m)
  speed_ms = 0.025
  movel([-0.015897, -0.699183, -2.792580, -1.220626, 1.570796, 1.554899],accel_mss,speed_ms,0,blend_radius_m)
  movel([-0.021119, -0.700059, -2.792469, -1.219861, 1.570796, 1.549677],accel_mss,speed_ms,0,blend_radius_m)
  movel([-0.023927, -0.700958, -2.792355, -1.219076, 1.570796, 1.546870],accel_mss,speed_ms,0,blend_radius_m)
  movel([-0.026870, -0.702245, -2.792191, -1.217953, 1.570796, 1.543926],accel_mss,speed_ms,0,blend_radius_m)
  movel([-0.029954, -0.703979, -2.791969, -1.216442, 1.570796, 1.540842],accel_mss,speed_ms,0,blend_radius_m)
  movel([-0.033189, -0.706214, -2.791680, -1.214494, 1.570796, 1.537607],accel_mss,speed_ms,0,blend_radius_m)
  speed_ms = 0.005
  movel([-0.033189, -0.699746, -2.785064, -1.227579, 1.570796, 1.537607],accel_mss,speed_ms,0,blend_radius_m)
  speed_ms = 0.040
  movel([-0.024336, -0.685951, -2.786799, -1.239639, 1.570796, 1.546460],accel_mss,speed_ms,0,blend_radius_m)
  speed_ms = 0.005
  movel([-0.024336, -0.692234, -2.793447, -1.226708, 1.570796, 1.546460],accel_mss,speed_ms,0,blend_radius_m)
  speed_ms = 0.025
  movel([-0.024945, -0.688308, -2.793927, -1.230154, 1.570796, 1.545851],accel_mss,speed_ms,0,blend_radius_m)
  movel([-0.026464, -0.685335, -2.794286, -1.232768, 1.570796, 1.544332],accel_mss,speed_ms,0,blend_radius_m)
  movel([-0.028811, -0.683327, -2.794526, -1.234536, 1.570796, 1.541985],accel_mss,speed_ms,0,blend_radius_m)
  movel([-0.031911, -0.682320, -2.794646, -1.235423, 1.570796, 1.538886],accel_mss,speed_ms,0,blend_radius_m)
  movel([-0.035676, -0.682328, -2.794645, -1.235416, 1.570796, 1.535120],accel_mss,speed_ms,0,blend_radius_m)
  movel([-0.040010, -0.683363, -2.794522, -1.234504, 1.570796, 1.530787],accel_mss,speed_ms,0,blend_radius_m)
  movel([-0.044815, -0.685428, -2.794275, -1.232686, 1.570796, 1.525981],accel_mss,speed_ms,0,blend_radius_m)
  movel([-0.047367, -0.686853, -2.794103, -1.231433, 1.570796, 1.523429],accel_mss,speed_ms,0,blend_radius_m)
  movel([-0.049997, -0.688527, -2.793900, -1.229962, 1.570796, 1.520799],accel_mss,speed_ms,0,blend_radius_m)
  speed_ms = 0.005
  movel([-0.049997, -0.682295, -2.787244, -1.242850, 1.570796, 1.520799],accel_mss,speed_ms,0,blend_radius_m)
  speed_ms = 0.040
  movel([-0.038264, -0.667878, -2.788942, -1.255570, 1.570796, 1.532533],accel_mss,speed_ms,0,blend_radius_m)
  speed_ms = 0.005
  movel([-0.038264, -0.673908, -2.795629, -1.242852, 1.570796, 1.532533],accel_mss,speed_ms,0,blend_radius_m)
  speed_ms = 0.025
  movel([-0.038980, -0.672328, -2.795810, -1.244251, 1.570796, 1.531816],accel_mss,speed_ms,0,blend_radius_m)
  movel([-0.039996, -0.671017, -2.795960, -1.245412, 1.570796, 1.530800],accel_mss,speed_ms,0,blend_radius_m)
  movel([-0.042840, -0.669199, -2.796166, -1.247025, 1.570796, 1.527956],accel_mss,speed_ms,0,blend_radius_m)
  movel([-0.046612, -0.668438, -2.796252, -1.247700, 1.570796, 1.524184],accel_mss,speed_ms,0,blend_radius_m)
  movel([-0.051114, -0.668716, -2.796220, -1.247453, 1.570796, 1.519683],accel_mss,speed_ms,0,blend_radius_m)
  movel([-0.056153, -0.669994, -2.796076, -1.246319, 1.570796, 1.514644],accel_mss,speed_ms,0,blend_radius_m)
  movel([-0.061509, -0.672222, -2.795822, -1.244345, 1.570796, 1.509288],accel_mss,speed_ms,0,blend_radius_m)
  movel([-0.064246, -0.673684, -2.795655, -1.243050, 1.570796, 1.506550],accel_mss,speed_ms,0,blend_radius_m)
  movel([-0.069697, -0.677252, -2.795242, -1.239895, 1.570796, 1.501099],accel_mss,speed_ms,0,blend_radius_m)
  movel([-0.072361, -0.679344, -2.794997, -1.238047, 1.570796, 1.498436],accel_mss,speed_ms,0,blend_radius_m)
  speed_ms = 0.005
  movel([-0.072361, -0.673238, -2.788321, -1.250829, 1.570796, 1.498436],accel_mss,speed_ms,0,blend_radius_m)
  speed_ms = 0.040
  movel([-0.055417, -0.654550, -2.790429, -1.267410, 1.570796, 1.515379],accel_mss,speed_ms,0,blend_radius_m)
  speed_ms = 0.005
  movel([-0.055417, -0.660388, -2.797144, -1.254857, 1.570796, 1.515379],accel_mss,speed_ms,0,blend_radius_m)
  speed_ms = 0.025
  movel([-0.059396, -0.659180, -2.797275, -1.255934, 1.570796, 1.511401],accel_mss,speed_ms,0,blend_radius_m)
  movel([-0.064045, -0.658961, -2.797299, -1.256129, 1.570796, 1.506751],accel_mss,speed_ms,0,blend_radius_m)
  movel([-0.069261, -0.659765, -2.797212, -1.255412, 1.570796, 1.501536],accel_mss,speed_ms,0,blend_radius_m)
  movel([-0.074961, -0.661610, -2.797010, -1.253769, 1.570796, 1.495836],accel_mss,speed_ms,0,blend_radius_m)
  movel([-0.081034, -0.664516, -2.796690, -1.251183, 1.570796, 1.489762],accel_mss,speed_ms,0,blend_radius_m)
  movel([-0.084180, -0.666367, -2.796484, -1.249538, 1.570796, 1.486617],accel_mss,speed_ms,0,blend_radius_m)
  movel([-0.087375, -0.668483, -2.796246, -1.247659, 1.570796, 1.483421],accel_mss,speed_ms,0,blend_radius_m)
  movel([-0.090616, -0.670871, -2.795976, -1.245542, 1.570796, 1.480180],accel_mss,speed_ms,0,blend_radius_m)
  movel([-0.093887, -0.673528, -2.795673, -1.243188, 1.570796, 1.476909],accel_mss,speed_ms,0,blend_radius_m)
  movel([-0.097168, -0.676446, -2.795336, -1.240607, 1.570796, 1.473628],accel_mss,speed_ms,0,blend_radius_m)
  movel([-0.100449, -0.679629, -2.794964, -1.237797, 1.570796, 1.470348],accel_mss,speed_ms,0,blend_radius_m)
  speed_ms = 0.005
  movel([-0.100449, -0.673519, -2.788289, -1.250582, 1.570796, 1.470348],accel_mss,speed_ms,0,blend_radius_m)
  speed_ms = 0.040
  movel([-0.083083, -0.651571, -2.790751, -1.270067, 1.570796, 1.487714],accel_mss,speed_ms,0,blend_radius_m)
  speed_ms = 0.005
  movel([-0.083083, -0.657366, -2.797472, -1.257551, 1.570796, 1.487714],accel_mss,speed_ms,0,blend_radius_m)
  speed_ms = 0.025
  movel([-0.084686, -0.655587, -2.797663, -1.259139, 1.570796, 1.486111],accel_mss,speed_ms,0,blend_radius_m)
  movel([-0.086796, -0.654423, -2.797787, -1.260179, 1.570796, 1.484000],accel_mss,speed_ms,0,blend_radius_m)
  movel([-0.089374, -0.653898, -2.797843, -1.260648, 1.570796, 1.481422],accel_mss,speed_ms,0,blend_radius_m)
  movel([-0.092367, -0.654029, -2.797829, -1.260531, 1.570796, 1.478429],accel_mss,speed_ms,0,blend_radius_m)
  movel([-0.096431, -0.655019, -2.797724, -1.259647, 1.570796, 1.474365],accel_mss,speed_ms,0,blend_radius_m)
  movel([-0.100822, -0.656708, -2.797543, -1.258139, 1.570796, 1.469975],accel_mss,speed_ms,0,blend_radius_m)
  movel([-0.106228, -0.659332, -2.797259, -1.255798, 1.570796, 1.464568],accel_mss,speed_ms,0,blend_radius_m)
  movel([-0.111818, -0.662625, -2.796899, -1.252865, 1.570796, 1.458979],accel_mss,speed_ms,0,blend_radius_m)
  movel([-0.117500, -0.666593, -2.796459, -1.249337, 1.570796, 1.453297],accel_mss,speed_ms,0,blend_radius_m)
  movel([-0.123186, -0.671251, -2.795933, -1.245205, 1.570796, 1.447611],accel_mss,speed_ms,0,blend_radius_m)
  movel([-0.128760, -0.676591, -2.795319, -1.240479, 1.570796, 1.442037],accel_mss,speed_ms,0,blend_radius_m)
  movel([-0.131440, -0.679473, -2.794982, -1.237934, 1.570796, 1.439356],accel_mss,speed_ms,0,blend_radius_m)
  movel([-0.136442, -0.685533, -2.794262, -1.232594, 1.570796, 1.434355],accel_mss,speed_ms,0,blend_radius_m)
  movel([-0.138714, -0.688661, -2.793884, -1.229844, 1.570796, 1.432082],accel_mss,speed_ms,0,blend_radius_m)
  movel([-0.140791, -0.691821, -2.793498, -1.227070, 1.570796, 1.430006],accel_mss,speed_ms,0,blend_radius_m)
  movel([-0.142651, -0.694993, -2.793105, -1.224290, 1.570796, 1.428145],accel_mss,speed_ms,0,blend_radius_m)
  speed_ms = 0.005
  movel([-0.142651, -0.688674, -2.786463, -1.237252, 1.570796, 1.428145],accel_mss,speed_ms,0,blend_radius_m)
  speed_ms = 0.040
  movel([-0.125872, -0.659959, -2.789835, -1.262595, 1.570796, 1.444924],accel_mss,speed_ms,0,blend_radius_m)
  speed_ms = 0.005
  movel([-0.125872, -0.665876, -2.796539, -1.249974, 1.570796, 1.444924],accel_mss,speed_ms,0,blend_radius_m)
  speed_ms = 0.025
  movel([-0.132879, -0.669628, -2.796117, -1.246644, 1.570796, 1.437918],accel_mss,speed_ms,0,blend_radius_m)
  movel([-0.140179, -0.674234, -2.795591, -1.242563, 1.570796, 1.430617],accel_mss,speed_ms,0,blend_radius_m)
  movel([-0.147568, -0.679639, -2.794963, -1.237787, 1.570796, 1.423228],accel_mss,speed_ms,0,blend_radius_m)
  movel([-0.151231, -0.682617, -2.794611, -1.235161, 1.570796, 1.419565],accel_mss,speed_ms,0,blend_radius_m)
  movel([-0.154841, -0.685772, -2.794233, -1.232383, 1.570796, 1.415955],accel_mss,speed_ms,0,blend_radius_m)
  movel([-0.158366, -0.689089, -2.793832, -1.229468, 1.570796, 1.412430],accel_mss,speed_ms,0,blend_radius_m)
  movel([-0.161780, -0.692556, -2.793407, -1.226426, 1.570796, 1.409016],accel_mss,speed_ms,0,blend_radius_m)
  movel([-0.165063, -0.696170, -2.792958, -1.223261, 1.570796, 1.405733],accel_mss,speed_ms,0,blend_radius_m)
  movel([-0.168188, -0.699923, -2.792486, -1.219980, 1.570796, 1.402608],accel_mss,speed_ms,0,blend_radius_m)
  movel([-0.171138, -0.703805, -2.791991, -1.216593, 1.570796, 1.399659],accel_mss,speed_ms,0,blend_radius_m)
  movel([-0.173875, -0.707804, -2.791474, -1.213111, 1.570796, 1.396921],accel_mss,speed_ms,0,blend_radius_m)
  movel([-0.176389, -0.711915, -2.790934, -1.209540, 1.570796, 1.394408],accel_mss,speed_ms,0,blend_radius_m)
  movel([-0.178649, -0.716130, -2.790373, -1.205886, 1.570796, 1.392148],accel_mss,speed_ms,0,blend_radius_m)
  speed_ms = 0.005
  movel([-0.178649, -0.709533, -2.783780, -1.219076, 1.570796, 1.392148],accel_mss,speed_ms,0,blend_radius_m)
  speed_ms = 0.040
  movel([-0.168864, -0.682306, -2.787243, -1.242840, 1.570796, 1.401933],accel_mss,speed_ms,0,blend_radius_m)
  speed_ms = 0.005
  movel([-0.168864, -0.688538, -2.793899, -1.229952, 1.570796, 1.401933],accel_mss,speed_ms,0,blend_radius_m)
  speed_ms = 0.025
  movel([-0.172372, -0.690671, -2.793639, -1.228080, 1.570796, 1.398424],accel_mss,speed_ms,0,blend_radius_m)
  movel([-0.175931, -0.693127, -2.793337, -1.225925, 1.570796, 1.394866],accel_mss,speed_ms,0,blend_radius_m)
  movel([-0.179494, -0.695880, -2.792995, -1.223515, 1.570796, 1.391302],accel_mss,speed_ms,0,blend_radius_m)
  movel([-0.183035, -0.698892, -2.792616, -1.220880, 1.570796, 1.387761],accel_mss,speed_ms,0,blend_radius_m)
  movel([-0.186523, -0.702140, -2.792204, -1.218045, 1.570796, 1.384273],accel_mss,speed_ms,0,blend_radius_m)
  movel([-0.189918, -0.705587, -2.791761, -1.215040, 1.570796, 1.380878],accel_mss,speed_ms,0,blend_radius_m)
  movel([-0.193188, -0.709198, -2.791292, -1.211899, 1.570796, 1.377608],accel_mss,speed_ms,0,blend_radius_m)
  movel([-0.196310, -0.712953, -2.790797, -1.208639, 1.570796, 1.374487],accel_mss,speed_ms,0,blend_radius_m)
  movel([-0.199241, -0.716811, -2.790281, -1.205297, 1.570796, 1.371555],accel_mss,speed_ms,0,blend_radius_m)
  movel([-0.201961, -0.720731, -2.789751, -1.201908, 1.570796, 1.368836],accel_mss,speed_ms,0,blend_radius_m)
  movel([-0.204448, -0.724673, -2.789210, -1.198506, 1.570796, 1.366348],accel_mss,speed_ms,0,blend_radius_m)
  movel([-0.206688, -0.728608, -2.788662, -1.195119, 1.570796, 1.364108],accel_mss,speed_ms,0,blend_radius_m)
  movel([-0.208668, -0.732499, -2.788114, -1.191776, 1.570796, 1.362128],accel_mss,speed_ms,0,blend_radius_m)
  movel([-0.210372, -0.736321, -2.787568, -1.188500, 1.570796, 1.360424],accel_mss,speed_ms,0,blend_radius_m)
  movel([-0.211774, -0.740026, -2.787032, -1.185331, 1.570796, 1.359023],accel_mss,speed_ms,0,blend_radius_m)
  movel([-0.212870, -0.743592, -2.786510, -1.182286, 1.570796, 1.357926],accel_mss,speed_ms,0,blend_radius_m)
  speed_ms = 0.005
  movel([-0.212870, -0.736656, -2.779984, -1.195748, 1.570796, 1.357926],accel_mss,speed_ms,0,blend_radius_m)
  speed_ms = 0.040
  movel([-0.209556, -0.714306, -2.783137, -1.214946, 1.570796, 1.361240],accel_mss,speed_ms,0,blend_radius_m)
  speed_ms = 0.005
  movel([-0.209556, -0.720964, -2.789719, -1.201706, 1.570796, 1.361240],accel_mss,speed_ms,0,blend_radius_m)
  speed_ms = 0.025
  movel([-0.212888, -0.723189, -2.789414, -1.199786, 1.570796, 1.357909],accel_mss,speed_ms,0,blend_radius_m)
  movel([-0.216197, -0.725887, -2.789041, -1.197460, 1.570796, 1.354599],accel_mss,speed_ms,0,blend_radius_m)
  movel([-0.219435, -0.728973, -2.788611, -1.194805, 1.570796, 1.351362],accel_mss,speed_ms,0,blend_radius_m)
  movel([-0.222573, -0.732364, -2.788133, -1.191892, 1.570796, 1.348223],accel_mss,speed_ms,0,blend_radius_m)
  movel([-0.225576, -0.735983, -2.787617, -1.188790, 1.570796, 1.345221],accel_mss,speed_ms,0,blend_radius_m)
  movel([-0.228402, -0.739743, -2.787073, -1.185573, 1.570796, 1.342394],accel_mss,speed_ms,0,blend_radius_m)
  movel([-0.231032, -0.743568, -2.786514, -1.182307, 1.570796, 1.339765],accel_mss,speed_ms,0,blend_radius_m)
  movel([-0.233420, -0.747379, -2.785949, -1.179061, 1.570796, 1.337376],accel_mss,speed_ms,0,blend_radius_m)
  movel([-0.235655, -0.751285, -2.785363, -1.175741, 1.570796, 1.335141],accel_mss,speed_ms,0,blend_radius_m)
  movel([-0.237660, -0.755173, -2.784772, -1.172444, 1.570796, 1.333137],accel_mss,speed_ms,0,blend_radius_m)
  movel([-0.239399, -0.758998, -2.784184, -1.169208, 1.570796, 1.331397],accel_mss,speed_ms,0,blend_radius_m)
  movel([-0.240817, -0.762693, -2.783608, -1.166088, 1.570796, 1.329979],accel_mss,speed_ms,0,blend_radius_m)
  movel([-0.241880, -0.766204, -2.783055, -1.163131, 1.570796, 1.328916],accel_mss,speed_ms,0,blend_radius_m)
  movel([-0.242547, -0.769478, -2.782533, -1.160377, 1.570796, 1.328249],accel_mss,speed_ms,0,blend_radius_m)
  movel([-0.242764, -0.772455, -2.782054, -1.157879, 1.570796, 1.328032],accel_mss,speed_ms,0,blend_radius_m)
  movel([-0.242503, -0.775088, -2.781627, -1.155674, 1.570796, 1.328293],accel_mss,speed_ms,0,blend_radius_m)
  speed_ms = 0.005
  movel([-0.242503, -0.767791, -2.775185, -1.169413, 1.570796, 1.328293],accel_mss,speed_ms,0,blend_radius_m)
  speed_ms = 0.040
  movel([-0.247417, -0.754226, -2.777335, -1.180828, 1.570796, 1.323380],accel_mss,speed_ms,0,blend_radius_m)
  speed_ms = 0.005
  movel([-0.247417, -0.761370, -2.783815, -1.167204, 1.570796, 1.323380],accel_mss,speed_ms,0,blend_radius_m)
  speed_ms = 0.025
  movel([-0.251512, -0.766168, -2.783060, -1.163160, 1.570796, 1.319284],accel_mss,speed_ms,0,blend_radius_m)
  movel([-0.255526, -0.771459, -2.782215, -1.158715, 1.570796, 1.315270],accel_mss,speed_ms,0,blend_radius_m)
  movel([-0.259229, -0.776987, -2.781317, -1.154085, 1.570796, 1.311567],accel_mss,speed_ms,0,blend_radius_m)
  movel([-0.262396, -0.782501, -2.780405, -1.149483, 1.570796, 1.308401],accel_mss,speed_ms,0,blend_radius_m)
  movel([-0.264815, -0.787767, -2.779520, -1.145102, 1.570796, 1.305981],accel_mss,speed_ms,0,blend_radius_m)
  movel([-0.265681, -0.790238, -2.779099, -1.143052, 1.570796, 1.305115],accel_mss,speed_ms,0,blend_radius_m)
  movel([-0.266280, -0.792556, -2.778702, -1.141131, 1.570796, 1.304516],accel_mss,speed_ms,0,blend_radius_m)
  movel([-0.266591, -0.794705, -2.778331, -1.139353, 1.570796, 1.304205],accel_mss,speed_ms,0,blend_radius_m)
  movel([-0.266590, -0.796654, -2.777993, -1.137742, 1.570796, 1.304206],accel_mss,speed_ms,0,blend_radius_m)
  movel([-0.266245, -0.798366, -2.777694, -1.136329, 1.570796, 1.304552],accel_mss,speed_ms,0,blend_radius_m)
  movel([-0.265537, -0.799831, -2.777437, -1.135121, 1.570796, 1.305260],accel_mss,speed_ms,0,blend_radius_m)
  speed_ms = 0.005
  movel([-0.265537, -0.792273, -2.771064, -1.149052, 1.570796, 1.305260],accel_mss,speed_ms,0,blend_radius_m)
  speed_ms = 0.040
  movel([-0.274720, -0.792530, -2.771019, -1.148840, 1.570796, 1.296076],accel_mss,speed_ms,0,blend_radius_m)
  speed_ms = 0.005
  movel([-0.274720, -0.800090, -2.777391, -1.134907, 1.570796, 1.296076],accel_mss,speed_ms,0,blend_radius_m)
  speed_ms = 0.025
  movel([-0.278738, -0.807730, -2.776031, -1.128628, 1.570796, 1.292058],accel_mss,speed_ms,0,blend_radius_m)
  movel([-0.280470, -0.811524, -2.775344, -1.125521, 1.570796, 1.290326],accel_mss,speed_ms,0,blend_radius_m)
  movel([-0.281915, -0.815203, -2.774670, -1.122516, 1.570796, 1.288882],accel_mss,speed_ms,0,blend_radius_m)
  movel([-0.282993, -0.818707, -2.774021, -1.119660, 1.570796, 1.287803],accel_mss,speed_ms,0,blend_radius_m)
  movel([-0.283636, -0.821978, -2.773410, -1.117001, 1.570796, 1.287160],accel_mss,speed_ms,0,blend_radius_m)
  movel([-0.283762, -0.824945, -2.772850, -1.114594, 1.570796, 1.287034],accel_mss,speed_ms,0,blend_radius_m)
  movel([-0.283305, -0.827559, -2.772353, -1.112477, 1.570796, 1.287491],accel_mss,speed_ms,0,blend_radius_m)
  speed_ms = 0.005
  # Splitting Linear movement in 2 (instruction 3386: MoveL 3110)
  movel([-0.283305, -0.808638, -2.756582, -1.147169, 1.570796, 1.287491],accel_mss,speed_ms,0,blend_radius_m)
  movel([-0.283305, -0.791754, -2.740670, -1.179965, 1.570796, 1.287491],accel_mss,speed_ms,0,blend_radius_m)
  speed_ms = 1.000
  movel([-0.283305, -0.791754, -2.740670, -1.179965, 1.570796, 1.287491],accel_mss,speed_ms,0,blend_radius_m)
  # Splitting Linear movement in 6 (instruction 3389: MoveL 3112)
  movel([-0.283305, -0.767608, -2.713865, -1.230916, 1.570796, 1.287491],accel_mss,speed_ms,0,blend_radius_m)
  movel([-0.283305, -0.747787, -2.686742, -1.277859, 1.570796, 1.287491],accel_mss,speed_ms,0,blend_radius_m)
  movel([-0.283305, -0.731650, -2.659333, -1.321406, 1.570796, 1.287491],accel_mss,speed_ms,0,blend_radius_m)
  movel([-0.283305, -0.718672, -2.631661, -1.362056, 1.570796, 1.287491],accel_mss,speed_ms,0,blend_radius_m)
  movel([-0.283305, -0.708419, -2.603744, -1.400226, 1.570796, 1.287491],accel_mss,speed_ms,0,blend_radius_m)
  movel([-0.283305, -0.700534, -2.575596, -1.436260, 1.570796, 1.287491],accel_mss,speed_ms,0,blend_radius_m)
  # End of main program
end

Machining1()
